// TIA Portal V21 export
// export: Created 2026-10-12T11:32:17.360201Z, ExportSetting WithDefaults, DisplayName Totally Integrated Automation Portal, DisplayVersion V21, DisplayName STEP 7 Professional, DisplayVersion V21, DisplayName STEP 7 Safety, DisplayVersion V21, DisplayName Tech WebApplication, DisplayVersion V21, DisplayName WinCC Basic/Comfort/Advanced, DisplayVersion V21, DisplayName WinCC Unified, DisplayVersion V21
VAR_GLOBAL   // PLC tag table "DI"
   "DI_PRODUCT SENSOR" AT %I0.0 : Bool;
   "DI_AUTO MANUAL SELECTION" AT %I0.1 : Bool;
   "DI_CYCLE START PB" AT %I0.2 : Bool;
   "DI_CYCLE STOP PB" AT %I0.3 : Bool;
   "DI_EMERGENCY PB" AT %I0.4 : Bool;
   "DI_CONVEYOR VFD FAULT" AT %I0.5 : Bool;
   "DI_SPARE I0.6" AT %I0.6 : Bool;
   "DI_SPARE I0.7" AT %I0.7 : Bool;
   "DI_SPARE I1.0" AT %I1.0 : Bool;
   "DI_SPARE I1.1" AT %I1.1 : Bool;
   "DI_SPARE I1.2" AT %I1.2 : Bool;
   "DI_SPARE I1.3" AT %I1.3 : Bool;
   "DI_SPARE I1.4" AT %I1.4 : Bool;
   "DI_SPARE I1.5" AT %I1.5 : Bool;
END_VAR
